// TIA Portal V19 export
TYPE "ST_Joggong"
   STRUCT
      Busy : Bool;
      Done : Bool;
      Error : Bool;
      "Error ID" : Word;
      FWD : Bool;
      BWD : Bool;
      Velocity : Real;
      Command_Aborted : Bool;
   END_STRUCT;
END_TYPE
